(* PLC project Vn_fb_user, Beckhoff Automation GmbH TwinCAT PLC Control 3.5.13.21 *)
(* stored: creationDateTime 1970-01-01T00:00:00 *)

PROGRAM Vn_fb_user

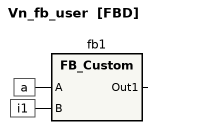
(* FBD diagram, written out as Structured Text *)
fb1(A := a, B := i1);
END_PROGRAM
